FUNCTION_BLOCK FB_FillingMarinade
VAR_INPUT
	iFillAmoungKg		: UINT;
	rActWeight			: REAL;
	bStop				: BOOL;
END_VAR
VAR_OUTPUT
	bFillingBusy		: BOOL;
	bFillingDone		: BOOL;
END_VAR
VAR_IN_OUT
	bFillRequest		: BOOL;
	fbFiliingPump		: FB_Pump;
	bPistonOpen			: BOOL;
	bPistonClose		: BOOL;
END_VAR
VAR
	trigStop			: R_TRIG;
	rHighVelocity		: REAL:=200;
	rMidVelocity		: REAL:=100;
	rLowVelocity		: REAL:=10;
END_VAR

actFillComponent();

trigStop(Clk:= bStop);
IF SFCReset THEN
	SFCReset:=FALSE;
END_IF
IF trigStop.Q THEN
	bFillRequest:=FALSE;
	SFCReset:=TRUE;
END_IF

ACTION actFillComponent:
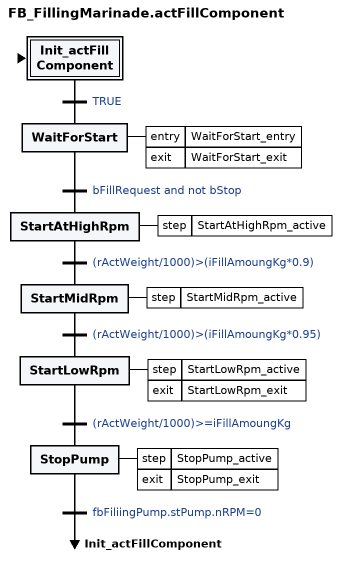
INITIAL_STEP Init_actFillComponent:
END_STEP
TRANSITION FROM Init_actFillComponent TO WaitForStart
    := TRUE;
END_TRANSITION
STEP WaitForStart:
    WaitForStart_entry(P1);  // entry action
    WaitForStart_exit(P0);  // exit action
END_STEP
TRANSITION FROM WaitForStart TO StartAtHighRpm
    := bFillRequest and not bStop;
END_TRANSITION
STEP StartAtHighRpm:
    StartAtHighRpm_active(N);  // step action
END_STEP
TRANSITION FROM StartAtHighRpm TO StartMidRpm
    := (rActWeight/1000)>(iFillAmoungKg*0.9);
END_TRANSITION
STEP StartMidRpm:
    StartMidRpm_active(N);  // step action
END_STEP
TRANSITION FROM StartMidRpm TO StartLowRpm
    := (rActWeight/1000)>(iFillAmoungKg*0.95);
END_TRANSITION
STEP StartLowRpm:
    StartLowRpm_active(N);  // step action
    StartLowRpm_exit(P0);  // exit action
END_STEP
TRANSITION FROM StartLowRpm TO StopPump
    := (rActWeight/1000)>=iFillAmoungKg;
END_TRANSITION
STEP StopPump:
    StopPump_active(N);  // step action
    StopPump_exit(P0);  // exit action
END_STEP
TRANSITION FROM StopPump TO Init_actFillComponent
    := fbFiliingPump.stPump.nRPM=0;
END_TRANSITION
END_ACTION

ACTION StartAtHighRpm_active:
fbFiliingPump.m_Run(RPM:=rHighVelocity);
END_ACTION

ACTION StartLowRpm_active:
fbFiliingPump.m_Run(RPM:=rMidVelocity);
END_ACTION

ACTION StartLowRpm_exit:
bPistonOpen:=FALSE;
bPistonClose:=TRUE;
END_ACTION

ACTION StartMidRpm_active:
fbFiliingPump.m_Run(RPM:=rMidVelocity);
END_ACTION

ACTION StopPump_active:
fbFiliingPump.m_Stop();
END_ACTION

ACTION StopPump_exit:
bFillingBusy:=FALSE;		
bFillingDone:=TRUE;
END_ACTION

ACTION WaitForStart_entry:
fbFiliingPump.m_Stop();
bPistonOpen:=FALSE;
bPistonClose:=TRUE;
END_ACTION

ACTION WaitForStart_exit:
bFillingBusy:=TRUE;		
bFillingDone:=FALSE;
bPistonOpen:=TRUE;
bPistonClose:=FALSE;
END_ACTION

END_FUNCTION_BLOCK

(* stored: Version 1.1.0.1, ProductVersion 3.1.4024.12
   POU FB_FillingMarinade: Id {e17c7fa9-00cf-4e3b-894a-a82205e0ff5f}, SpecialFunc None
   Folder Management: Id {2e571a8a-32c1-4b64-83bc-f923998c1f7e}
   Action actFillComponent: Id {6894fc14-c166-47b6-a362-77a3604bf65a}
   Action StartAtHighRpm_active: Id {bcded3d3-2299-4c62-a9f4-e9f8fe45261d}
   Action StartLowRpm_active: Id {380b44ce-b1e0-415e-8f91-c44e5a8f6dbc}
   Action StartLowRpm_exit: Id {2675f051-70de-4ef8-9c8e-4fc745d473b2}
   Action StartMidRpm_active: Id {bed15719-e5ab-41fa-8c93-5847edacd90c}
   Action StopPump_active: Id {e1e2b1da-bdbd-4bd0-99ba-c0c76a589a08}
   Action StopPump_exit: Id {2f39c003-3af6-4b1f-ae2a-096aade5d88f}
   Action WaitForStart_entry: Id {c6794e7c-ee45-4675-a817-40ea0922288e}
   Action WaitForStart_exit: Id {4d81a8f3-eaae-48f0-a92d-b9bcb5ae0c35} *)
